FUNCTION_BLOCK FB_LocalIntegrationTests EXTENDS TcUnit.FB_TestSuite
VAR
END_VAR

MappingInputs();
MappingOutputs();
FullChain();
HallSimulationChain();

METHOD PRIVATE MappingInputs
VAR
    fbInputs : FB_SimulationInputs;
    bWorkshopButton : BOOL;
    bEntrywayLowerButton : BOOL;
    bEntrywayUpperButton : BOOL;
    stInputs : ST_HomeInputs;
END_VAR
TEST('Simulation inputs map all button fields');

bWorkshopButton := FALSE;
bEntrywayLowerButton := FALSE;
bEntrywayUpperButton := FALSE;
fbInputs(
    bWorkshopButton := bWorkshopButton,
    bEntrywayLowerButton := bEntrywayLowerButton,
    bEntrywayUpperButton := bEntrywayUpperButton,
    stInputs => stInputs);
AssertTrue(Condition := NOT stInputs.Workshop.bButton, Message := 'Workshop button maps low');
AssertTrue(Condition := NOT stInputs.Entryway.bLowerButton, Message := 'Entryway button maps low');
AssertTrue(Condition := NOT stInputs.Entryway.bUpperButton, Message := 'Entryway upper button maps low');

bWorkshopButton := TRUE;
fbInputs(
    bWorkshopButton := bWorkshopButton,
    bEntrywayLowerButton := bEntrywayLowerButton,
    bEntrywayUpperButton := bEntrywayUpperButton,
    stInputs => stInputs);
AssertTrue(Condition := stInputs.Workshop.bButton, Message := 'Workshop button maps high');
AssertTrue(Condition := NOT stInputs.Entryway.bLowerButton, Message := 'Entryway button remains low');
AssertTrue(Condition := NOT stInputs.Entryway.bUpperButton, Message := 'Entryway upper button remains low');

bWorkshopButton := FALSE;
bEntrywayLowerButton := TRUE;
fbInputs(
    bWorkshopButton := bWorkshopButton,
    bEntrywayLowerButton := bEntrywayLowerButton,
    bEntrywayUpperButton := bEntrywayUpperButton,
    stInputs => stInputs);
AssertTrue(Condition := NOT stInputs.Workshop.bButton, Message := 'Workshop button remains low');
AssertTrue(Condition := stInputs.Entryway.bLowerButton, Message := 'Entryway button maps high');
AssertTrue(Condition := NOT stInputs.Entryway.bUpperButton, Message := 'Entryway upper button remains low');

bEntrywayLowerButton := FALSE;
bEntrywayUpperButton := TRUE;
fbInputs(
    bWorkshopButton := bWorkshopButton,
    bEntrywayLowerButton := bEntrywayLowerButton,
    bEntrywayUpperButton := bEntrywayUpperButton,
    stInputs => stInputs);
AssertTrue(Condition := NOT stInputs.Workshop.bButton, Message := 'Workshop button remains low');
AssertTrue(Condition := NOT stInputs.Entryway.bLowerButton, Message := 'Entryway button remains low');
AssertTrue(Condition := stInputs.Entryway.bUpperButton, Message := 'Entryway upper button maps high');

TEST_FINISHED();
END_METHOD

METHOD PRIVATE MappingOutputs
VAR
    fbOutputs : FB_SimulationOutputs;
    stOutputs : ST_HomeOutputs;
    bWorkshopLightRelay : BOOL;
    bEntrywayLightRelay : BOOL;
    bEntrywayTemporaryLightRelay : BOOL;
    bHallOuterSpotsRelay : BOOL;
    bHallMiddleSpotRelay : BOOL;
END_VAR
TEST('Simulation outputs map all relay fields');

bWorkshopLightRelay := TRUE;
bEntrywayLightRelay := TRUE;
bEntrywayTemporaryLightRelay := TRUE;
bHallOuterSpotsRelay := TRUE;
bHallMiddleSpotRelay := TRUE;
stOutputs.Workshop.bLightRelay := FALSE;
stOutputs.Entryway.bLightRelay := FALSE;
stOutputs.Entryway.bTemporaryLightRelay := FALSE;
stOutputs.Hall.bOuterSpotsRelay := FALSE;
stOutputs.Hall.bMiddleSpotRelay := FALSE;
fbOutputs(
    stOutputs := stOutputs,
    bWorkshopLightRelay := bWorkshopLightRelay,
    bEntrywayLightRelay := bEntrywayLightRelay,
    bEntrywayTemporaryLightRelay := bEntrywayTemporaryLightRelay,
    bHallOuterSpotsRelay := bHallOuterSpotsRelay,
    bHallMiddleSpotRelay := bHallMiddleSpotRelay);
AssertTrue(Condition := NOT bWorkshopLightRelay, Message := 'Workshop relay maps low');
AssertTrue(Condition := NOT bEntrywayLightRelay, Message := 'Entryway relay maps low');
AssertTrue(Condition := NOT bEntrywayTemporaryLightRelay, Message := 'Entryway temporary relay maps low');

stOutputs.Workshop.bLightRelay := TRUE;
fbOutputs(
    stOutputs := stOutputs,
    bWorkshopLightRelay := bWorkshopLightRelay,
    bEntrywayLightRelay := bEntrywayLightRelay,
    bEntrywayTemporaryLightRelay := bEntrywayTemporaryLightRelay,
    bHallOuterSpotsRelay := bHallOuterSpotsRelay,
    bHallMiddleSpotRelay := bHallMiddleSpotRelay);
AssertTrue(Condition := bWorkshopLightRelay, Message := 'Workshop relay maps high');
AssertTrue(Condition := NOT bEntrywayLightRelay, Message := 'Entryway relay remains low');
AssertTrue(Condition := NOT bEntrywayTemporaryLightRelay, Message := 'Entryway temporary relay remains low');

stOutputs.Workshop.bLightRelay := FALSE;
stOutputs.Entryway.bLightRelay := TRUE;
fbOutputs(
    stOutputs := stOutputs,
    bWorkshopLightRelay := bWorkshopLightRelay,
    bEntrywayLightRelay := bEntrywayLightRelay,
    bEntrywayTemporaryLightRelay := bEntrywayTemporaryLightRelay,
    bHallOuterSpotsRelay := bHallOuterSpotsRelay,
    bHallMiddleSpotRelay := bHallMiddleSpotRelay);
AssertTrue(Condition := NOT bWorkshopLightRelay, Message := 'Workshop relay remains low');
AssertTrue(Condition := bEntrywayLightRelay, Message := 'Entryway relay maps high');
AssertTrue(Condition := NOT bEntrywayTemporaryLightRelay, Message := 'Entryway temporary relay remains low');

stOutputs.Entryway.bLightRelay := FALSE;
stOutputs.Entryway.bTemporaryLightRelay := TRUE;
fbOutputs(
    stOutputs := stOutputs,
    bWorkshopLightRelay := bWorkshopLightRelay,
    bEntrywayLightRelay := bEntrywayLightRelay,
    bEntrywayTemporaryLightRelay := bEntrywayTemporaryLightRelay,
    bHallOuterSpotsRelay := bHallOuterSpotsRelay,
    bHallMiddleSpotRelay := bHallMiddleSpotRelay);
AssertTrue(Condition := NOT bWorkshopLightRelay, Message := 'Workshop relay remains low');
AssertTrue(Condition := NOT bEntrywayLightRelay, Message := 'Entryway relay remains low');
AssertTrue(Condition := bEntrywayTemporaryLightRelay, Message := 'Entryway temporary relay maps high');

stOutputs.Entryway.bTemporaryLightRelay := FALSE;
fbOutputs(
    stOutputs := stOutputs,
    bWorkshopLightRelay := bWorkshopLightRelay,
    bEntrywayLightRelay := bEntrywayLightRelay,
    bEntrywayTemporaryLightRelay := bEntrywayTemporaryLightRelay,
    bHallOuterSpotsRelay := bHallOuterSpotsRelay,
    bHallMiddleSpotRelay := bHallMiddleSpotRelay);
AssertTrue(Condition := NOT bWorkshopLightRelay, Message := 'Workshop relay maps low again');
AssertTrue(Condition := NOT bEntrywayLightRelay, Message := 'Entryway relay maps low again');
AssertTrue(Condition := NOT bEntrywayTemporaryLightRelay, Message := 'Entryway temporary relay maps low again');

TEST_FINISHED();
END_METHOD

METHOD PRIVATE FullChain
VAR
    fbInputs : FB_SimulationInputs;
    fbHome : FB_Home;
    fbOutputs : FB_SimulationOutputs;
    stInputs : ST_HomeInputs;
    stOutputs : ST_HomeOutputs;
    bWorkshopButton : BOOL;
    bEntrywayLowerButton : BOOL;
    bEntrywayUpperButton : BOOL;
    bWorkshopLightRelay : BOOL;
    bEntrywayLightRelay : BOOL;
    bEntrywayTemporaryLightRelay : BOOL;
    bHallOuterSpotsRelay : BOOL;
    bHallMiddleSpotRelay : BOOL;
    bExpectedWorkshopRelay : BOOL;
    bExpectedEntrywayRelay : BOOL;
    bExpectedEntrywayTemporaryRelay : BOOL;
    nCircuit : INT;
    nStep : INT;
END_VAR
TEST('Private simulation adapters run each relay circuit through Core');

bWorkshopLightRelay := TRUE;
bEntrywayLightRelay := TRUE;
bEntrywayTemporaryLightRelay := TRUE;
bHallOuterSpotsRelay := TRUE;
bHallMiddleSpotRelay := TRUE;

FOR nCircuit := 1 TO 3 DO
    FOR nStep := 0 TO 4 DO
        bWorkshopButton := FALSE;
        bEntrywayLowerButton := FALSE;
        bEntrywayUpperButton := FALSE;

        IF (nStep = 1) OR (nStep = 3) THEN
            CASE nCircuit OF
                1: bWorkshopButton := TRUE;
                2: bEntrywayLowerButton := TRUE;
                3: bEntrywayUpperButton := TRUE;
            END_CASE;
        END_IF;

        bExpectedWorkshopRelay := (nCircuit = 1) AND ((nStep = 1) OR (nStep = 2));
        bExpectedEntrywayRelay := (nCircuit = 2) AND ((nStep = 1) OR (nStep = 2));
        bExpectedEntrywayTemporaryRelay := (nCircuit = 3) AND ((nStep = 1) OR (nStep = 2));

        fbInputs(
            bWorkshopButton := bWorkshopButton,
            bEntrywayLowerButton := bEntrywayLowerButton,
            bEntrywayUpperButton := bEntrywayUpperButton,
            stInputs => stInputs);
        fbHome(stInputs := stInputs, stOutputs => stOutputs);
        fbOutputs(
            stOutputs := stOutputs,
            bWorkshopLightRelay := bWorkshopLightRelay,
            bEntrywayLightRelay := bEntrywayLightRelay,
            bEntrywayTemporaryLightRelay := bEntrywayTemporaryLightRelay,
            bHallOuterSpotsRelay := bHallOuterSpotsRelay,
            bHallMiddleSpotRelay := bHallMiddleSpotRelay);

        AssertTrue(Condition := stOutputs.Workshop.bLightRelay = bExpectedWorkshopRelay, Message := 'Core workshop relay follows its button sequence');
        AssertTrue(Condition := stOutputs.Entryway.bLightRelay = bExpectedEntrywayRelay, Message := 'Core entryway relay follows its button sequence');
        AssertTrue(Condition := stOutputs.Entryway.bTemporaryLightRelay = bExpectedEntrywayTemporaryRelay, Message := 'Core entryway temporary relay follows its button sequence');
        AssertTrue(Condition := bWorkshopLightRelay = bExpectedWorkshopRelay, Message := 'Workshop relay reaches private endpoint');
        AssertTrue(Condition := bEntrywayLightRelay = bExpectedEntrywayRelay, Message := 'Entryway relay reaches private endpoint');
        AssertTrue(Condition := bEntrywayTemporaryLightRelay = bExpectedEntrywayTemporaryRelay, Message := 'Entryway temporary relay reaches private endpoint');
    END_FOR;
END_FOR;

TEST_FINISHED();
END_METHOD

METHOD PRIVATE HallSimulationChain
VAR
    fbInputs : FB_SimulationInputs;
    fbOutputs : FB_SimulationOutputs;
    fbHome : FB_Home;
    stInputs : ST_HomeInputs;
    stOutputs : ST_HomeOutputs;
    bHallUpperButton : BOOL;
    bHallLowerButton : BOOL;
    bWorkshopLightRelay : BOOL;
    bEntrywayLightRelay : BOOL;
    bEntrywayTemporaryLightRelay : BOOL;
    bHallOuterSpotsRelay : BOOL;
    bHallMiddleSpotRelay : BOOL;
END_VAR
TEST('Hall simulation adapters propagate private inputs through Core to private relay endpoints');

bHallUpperButton := FALSE;
bHallLowerButton := FALSE;
fbInputs(
    bWorkshopButton := FALSE,
    bEntrywayLowerButton := FALSE,
    bEntrywayUpperButton := FALSE,
    bHallUpperButton := bHallUpperButton,
    bHallLowerButton := bHallLowerButton,
    stInputs => stInputs);
fbHome(stInputs := stInputs, stOutputs => stOutputs);
fbOutputs(
    stOutputs := stOutputs,
    bWorkshopLightRelay := bWorkshopLightRelay,
    bEntrywayLightRelay := bEntrywayLightRelay,
    bEntrywayTemporaryLightRelay := bEntrywayTemporaryLightRelay,
    bHallOuterSpotsRelay := bHallOuterSpotsRelay,
    bHallMiddleSpotRelay := bHallMiddleSpotRelay);

bHallLowerButton := TRUE;
fbInputs(
    bWorkshopButton := FALSE,
    bEntrywayLowerButton := FALSE,
    bEntrywayUpperButton := FALSE,
    bHallUpperButton := bHallUpperButton,
    bHallLowerButton := bHallLowerButton,
    stInputs => stInputs);
fbHome(stInputs := stInputs, stOutputs => stOutputs);
fbOutputs(
    stOutputs := stOutputs,
    bWorkshopLightRelay := bWorkshopLightRelay,
    bEntrywayLightRelay := bEntrywayLightRelay,
    bEntrywayTemporaryLightRelay := bEntrywayTemporaryLightRelay,
    bHallOuterSpotsRelay := bHallOuterSpotsRelay,
    bHallMiddleSpotRelay := bHallMiddleSpotRelay);
AssertTrue(Condition := bEntrywayLightRelay, Message := 'Hall lower button reaches private Entryway endpoint');

bHallLowerButton := FALSE;
bHallUpperButton := TRUE;
fbInputs(
    bWorkshopButton := FALSE,
    bEntrywayLowerButton := FALSE,
    bEntrywayUpperButton := FALSE,
    bHallUpperButton := bHallUpperButton,
    bHallLowerButton := bHallLowerButton,
    stInputs => stInputs);
fbHome(stInputs := stInputs, stOutputs => stOutputs);
fbOutputs(
    stOutputs := stOutputs,
    bWorkshopLightRelay := bWorkshopLightRelay,
    bEntrywayLightRelay := bEntrywayLightRelay,
    bEntrywayTemporaryLightRelay := bEntrywayTemporaryLightRelay,
    bHallOuterSpotsRelay := bHallOuterSpotsRelay,
    bHallMiddleSpotRelay := bHallMiddleSpotRelay);
AssertTrue(Condition := bHallOuterSpotsRelay AND bHallMiddleSpotRelay, Message := 'Hall upper reaches both private spot endpoints');
AssertTrue(Condition := bEntrywayLightRelay, Message := 'Hall upper leaves Entryway endpoint unchanged');

TEST_FINISHED();
END_METHOD

END_FUNCTION_BLOCK

(* stored: Version 1.1.0.1
   POU FB_LocalIntegrationTests: Id {E0C05F45-7AF9-4D8D-97C2-45DFD62AC86A}, SpecialFunc None
   Method MappingInputs: Id {0F2458A0-E5CC-483B-81E8-0485F0595D09}
   Method MappingOutputs: Id {EDECD1D8-51AB-4B8F-94E6-30B39F9A4DA7}
   Method FullChain: Id {8117CC6D-4996-4E4E-A573-D0B92951EB4C}
   Method HallSimulationChain: Id {be317531-6179-493c-a99d-716513c74d78} *)
